Fanuc KAREL source: kb00031.KL

-- PROVISIONAL review KL for V940-1; original PC SHA256 d3c17cccaa8a71d1bcd9bc8a785bfbc579af165ef97a8bd55959972e123186df
-- Incomplete behavior may be omitted. Consult companion uncertainty JSON. Do not deploy.
PROGRAM KB00031
%NOLOCKGROUP
BEGIN
  -- V9_ZERO_TABLE_METADATA_HINT layout=0002_ascii; no indexed target words; source/name/runtime held
  -- UNRESOLVED_PC offsets 5-16; opcodes 2E,23
  -- UNRESOLVED_PC offsets 21-30; opcodes 3F,75
  -- UNRESOLVED_PC offsets 35-42; opcodes 9D,23
  -- UNRESOLVED_PC offsets 47-71; opcodes 27,22,22,2A,22,31
  -- UNRESOLVED_PC offsets 76-80; opcodes 7F
END KB00031
